FUNCTION_BLOCK T_SafePulse_UserFB EXTENDS T_SafeFunctionBlockBase
VAR_INPUT
	TonIn1 : BOOL;
	Parameters : ST_SafeTimerParameters;
END_VAR
VAR_OUTPUT
	TonOut : BOOL;
END_VAR
VAR
	safeTon : T_SafeTon(_group);
	safeAnd : T_SafeAnd(_group);
END_VAR

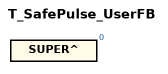
SUPER^();

METHOD FB_init : BOOL
VAR_INPUT
	bInitRetains	: BOOL;
	bInCopyCode	: BOOL;
	group	: REFERENCE TO T_SafeGroup;
END_VAR
safeAnd.SetGroupReference(bInCopyCode := bInCopyCode, group := group);
safeTon.SetGroupReference(bInCopyCode := bInCopyCode, group := group);
END_METHOD

METHOD PROTECTED Process
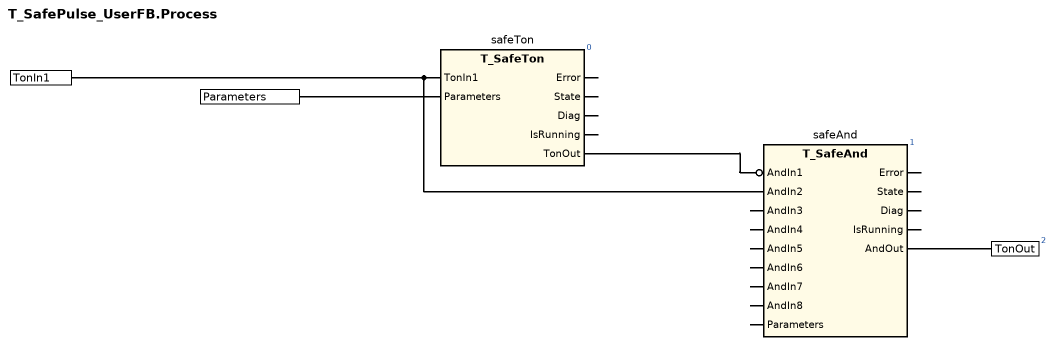
safeTon(TonIn1 := TonIn1, Parameters := Parameters); // T_SafeTon
safeAnd(AndIn1 := NOT safeTon.TonOut, AndIn2 := TonIn1); // T_SafeAnd
TonOut := safeAnd.AndOut;
END_METHOD

END_FUNCTION_BLOCK

(* stored: Version 1.1.0.1
   POU T_SafePulse_UserFB: Id {54b50892-fdaf-4337-b459-8dbdb773dd39}, SpecialFunc None
   Method FB_init: Id {a6f1625c-3374-4203-bef4-cd16712beb82}
   Method Process: Id {0fb23210-e247-4edb-afe7-513aa7d3aad4} *)
